(* IEC 61131-3 sources: repolevel_ST_code_completion/ground_truth/repoeval_modbus/readful_result, 6 files *)

(* ---- DataReverse_cmdReverse.st ---- *)
It seems like you are sharing code fragments from a repository, and you are particularly interested in the `cmdReverse` function and its context. However, the code snippet you provided at the end is incomplete. Let me help you understand the `cmdReverse` function and its purpose based on the fragments you have shared.

### `cmdReverse` Function Overview
The `cmdReverse` function is a simple function that takes an input of type `TargetDirect` and returns a `TargetDirect` value. The purpose of this function is to reverse the direction of a target. Based on the input value (`TargetDirect.extend` or `TargetDirect.retract`), it returns the opposite direction.

Here is the complete code for the `cmdReverse` function from the first fragment:

```pascal
FUNCTION cmdReverse : TargetDirect
VAR_INPUT
	input		:TargetDirect;
END_VAR

IF input = TargetDirect.extend THEN
	cmdReverse := TargetDirect.retract;
END_IF
IF input = TargetDirect.retract THEN
	cmdReverse := TargetDirect.extend;
END_IF
```

### Explanation
1. **Input Parameter**:
   - `input`: A variable of type `TargetDirect`, which presumably has two possible values: `extend` and `retract`.

2. **Logic**:
   - If the input is `TargetDirect.extend`, the function returns `TargetDirect.retract`.
   - If the input is `TargetDirect.retract`, the function returns `TargetDirect.extend`.

3. **Output**:
   - The function returns the reversed direction as a value of type `TargetDirect`.

### Usage Context
From the other fragments, it seems like this function is part of a larger system that involves Modbus communication and data handling. The `cmdReverse` function might be used in scenarios where the system needs to toggle or reverse the direction of a target, such as a motor or actuator.

For example:
- In the `localCmdHandler` method, variables like `exDirect` and `exeDirect` of type `TargetDirect` are declared. These might be used in conjunction with the `cmdReverse` function to handle commands that involve reversing directions.

### Missing Code
The last part of your message seems to repeat the `cmdReverse` function declaration but does not provide additional context or code. If you have specific questions or need further clarification, feel free to provide more details or ask!

(* ---- DataReverse_cmdReverse_1.st ---- *)
It seems like you are sharing code fragments from a repository, and you are particularly interested in the `cmdReverse` function and its context. However, the code snippet you provided at the end is incomplete. Let me help you understand the `cmdReverse` function and its purpose based on the fragments you have shared.

### `cmdReverse` Function Overview
The `cmdReverse` function is a simple function that takes an input of type `TargetDirect` and returns a `TargetDirect` value. The purpose of this function is to reverse the direction of a target. Based on the input value (`TargetDirect.extend` or `TargetDirect.retract`), it returns the opposite direction.

Here is the complete code for the `cmdReverse` function from the first fragment:

```pascal
FUNCTION cmdReverse : TargetDirect
VAR_INPUT
	input		:TargetDirect;
END_VAR

IF input = TargetDirect.extend THEN
	cmdReverse := TargetDirect.retract;
END_IF
IF input = TargetDirect.retract THEN
	cmdReverse := TargetDirect.extend;
END_IF
```

### Explanation
1. **Input Parameter**:
   - `input`: A variable of type `TargetDirect`, which presumably has two possible values: `extend` and `retract`.

2. **Logic**:
   - If the input is `TargetDirect.extend`, the function returns `TargetDirect.retract`.
   - If the input is `TargetDirect.retract`, the function returns `TargetDirect.extend`.

3. **Output**:
   - The function returns the reversed direction as a value of type `TargetDirect`.

### Usage Context
From the other fragments, it seems like this function is part of a larger system that involves Modbus communication and data handling. The `cmdReverse` function might be used in scenarios where the system needs to toggle or reverse the direction of a target, such as a motor or actuator.

For example:
- In the `localCmdHandler` method, variables like `exDirect` and `exeDirect` of type `TargetDirect` are declared. These might be used in conjunction with the `cmdReverse` function to handle commands that involve reversing directions.

### Missing Code
The last part of your message seems to repeat the `cmdReverse` function declaration but does not provide additional context or code. If you have specific questions or need further clarification, feel free to provide more details or ask!

(* ---- setButtonByDirect.st ---- *)
The provided code fragments define a function named `setButtonByDirect` in Structured Text (ST), which is commonly used in PLC programming. This function is designed to manipulate UI button variables based on input parameters such as `level`, `idx`, and `direct`.

### Function Overview:
- **Inputs:**
  - `level`: An integer indicating the type of track (1 for 地轨, 2 for 天轨).
  - `idx`: An integer representing the index of the挡板 (barrier).
  - `direct`: A variable of type `TargetDirect` that specifies the direction (`extend`, `retract`, or `stop`).

- **Purpose:**
  The function updates the state of UI button variables (`btnStop`, `btnExtend`, `btnRetract`) based on the input parameters.

### Key Observations:
1. **Parameter Validation:**
   - For `level = 1`, the function checks if `idx` is 0 or greater than 10. If this condition is true, the function exits early (`RETURN`).
   - For `level = 2`, the function checks if `idx` is greater than 10 and exits early if the condition is true.

2. **Button State Updates:**
   - Depending on the value of `direct` (`TargetDirect.extend`, `TargetDirect.retract`, or `TargetDirect.stop`), the function updates the button states (`btnStop`, `btnExtend`, `btnRetract`) for the specified `idx` in the `gUI.grd` array.

3. **Incomplete Code:**
   - The code fragments provided are incomplete. For example, the logic for `level = 2` is partially shown, and the handling of `TargetDirect.extend` for `level = 2` is missing.

### Suggestions for Improvement:
1. **Complete the Logic for `level = 2`:**
   - Ensure that all cases for `direct` (`extend`, `retract`, `stop`) are handled for `level = 2`.

2. **Add Comments for Clarity:**
   - While the code includes some comments, additional explanations for the logic (e.g., why certain conditions are checked) would improve readability.

3. **Error Handling:**
   - Consider adding error handling or logging for invalid input values to make debugging easier.

4. **Code Duplication:**
   - The logic for updating button states (`btnStop`, `btnExtend`, `btnRetract`) is duplicated for `level = 1` and `level = 2`. This could be refactored into a helper function to reduce redundancy.

### Example of Refactored Code:
```st
FUNCTION setButtonByDirect : BOOL
VAR_INPUT
	level		:INT;	// 1->地轨, 2->天轨
	idx			:INT;	// 挡板索引编号
	direct		:TargetDirect; // Direction
END_VAR
VAR
END_VAR

// Helper function to update button states
FUNCTION UpdateButtonStates : VOID
VAR_INPUT
	idx			:INT;
	direct		:TargetDirect;
END_VAR
BEGIN
	CASE direct OF
		TargetDirect.extend:
			gUI.grd[idx].btnStop := FALSE;
			gUI.grd[idx].btnExtend := TRUE;
			gUI.grd[idx].btnRetract := FALSE;
		TargetDirect.retract:
			gUI.grd[idx].btnStop := FALSE;
			gUI.grd[idx].btnExtend := FALSE;
			gUI.grd[idx].btnRetract := TRUE;
		TargetDirect.stop:
			gUI.grd[idx].btnStop := FALSE;
			gUI.grd[idx].btnExtend := FALSE;
			gUI.grd[idx].btnRetract := FALSE;
	END_CASE
END_FUNCTION

// Main function logic
BEGIN
	CASE level OF
		1:
			IF idx = 0 OR idx > 10 THEN
				RETURN;
			END_IF
			UpdateButtonStates(idx, direct);
		2:
			IF idx > 10 THEN
				RETURN;
			END_IF
			UpdateButtonStates(idx, direct);
	END_CASE
END_FUNCTION
```

This refactored version introduces a helper function `UpdateButtonStates` to handle button state updates, reducing code duplication and improving maintainability.

(* ---- setButtonByDirect_1.st ---- *)
The provided code fragments define a function named `setButtonByDirect` in Structured Text (ST), which is commonly used in PLC programming. This function is designed to manipulate UI button variables based on input parameters such as `level`, `idx`, and `direct`.

### Function Overview:
- **Inputs:**
  - `level`: An integer indicating the type of track (1 for 地轨, 2 for 天轨).
  - `idx`: An integer representing the index of the挡板 (barrier).
  - `direct`: A variable of type `TargetDirect` that specifies the direction (`extend`, `retract`, or `stop`).

- **Purpose:**
  The function updates the state of UI button variables (`btnStop`, `btnExtend`, `btnRetract`) based on the input parameters.

### Key Observations:
1. **Parameter Validation:**
   - For `level = 1`, the function checks if `idx` is 0 or greater than 10. If this condition is true, the function exits early (`RETURN`).
   - For `level = 2`, the function checks if `idx` is greater than 10 and exits early if the condition is true.

2. **Button State Updates:**
   - Depending on the value of `direct` (`TargetDirect.extend`, `TargetDirect.retract`, or `TargetDirect.stop`), the function updates the button states (`btnStop`, `btnExtend`, `btnRetract`) for the specified `idx` in the `gUI.grd` array.

3. **Incomplete Code:**
   - The code fragments provided are incomplete. For example, the logic for `level = 2` is partially shown, and the handling of `TargetDirect.extend` for `level = 2` is missing.

### Suggestions for Improvement:
1. **Complete the Logic for `level = 2`:**
   - Ensure that all cases for `direct` (`extend`, `retract`, `stop`) are handled for `level = 2`.

2. **Add Comments for Clarity:**
   - While the code includes some comments, additional explanations for the logic (e.g., why certain conditions are checked) would improve readability.

3. **Error Handling:**
   - Consider adding error handling or logging for invalid input values to make debugging easier.

4. **Code Duplication:**
   - The logic for updating button states (`btnStop`, `btnExtend`, `btnRetract`) is duplicated for `level = 1` and `level = 2`. This could be refactored into a helper function to reduce redundancy.

### Example of Refactored Code:
```st
FUNCTION setButtonByDirect : BOOL
VAR_INPUT
	level		:INT;	// 1->地轨, 2->天轨
	idx			:INT;	// 挡板索引编号
	direct		:TargetDirect; // Direction
END_VAR
VAR
END_VAR

// Helper function to update button states
FUNCTION UpdateButtonStates : VOID
VAR_INPUT
	idx			:INT;
	direct		:TargetDirect;
END_VAR
BEGIN
	CASE direct OF
		TargetDirect.extend:
			gUI.grd[idx].btnStop := FALSE;
			gUI.grd[idx].btnExtend := TRUE;
			gUI.grd[idx].btnRetract := FALSE;
		TargetDirect.retract:
			gUI.grd[idx].btnStop := FALSE;
			gUI.grd[idx].btnExtend := FALSE;
			gUI.grd[idx].btnRetract := TRUE;
		TargetDirect.stop:
			gUI.grd[idx].btnStop := FALSE;
			gUI.grd[idx].btnExtend := FALSE;
			gUI.grd[idx].btnRetract := FALSE;
	END_CASE
END_FUNCTION

// Main function logic
BEGIN
	CASE level OF
		1:
			IF idx = 0 OR idx > 10 THEN
				RETURN;
			END_IF
			UpdateButtonStates(idx, direct);
		2:
			IF idx > 10 THEN
				RETURN;
			END_IF
			UpdateButtonStates(idx, direct);
	END_CASE
END_FUNCTION
```

This refactored version introduces a helper function `UpdateButtonStates` to handle button state updates, reducing code duplication and improving maintainability.

(* ---- mdbsNumToIdx.st ---- *)
It seems like you are sharing multiple versions of a code fragment for a function block named `mdbsNumToIdx`. This function block takes a `devNo` (device number) as input and outputs `level` and `idx` based on the value of `devNo`. The code appears to be evolving across the fragments, with additional cases being added in each version.

Here’s a summary of the functionality and changes across the fragments:

---

### **Functionality**
1. **Input**:
   - `devNo`: A `WORD` (16-bit unsigned integer) representing the device number.

2. **Output**:
   - `level`: An `INT` (integer) representing the level associated with the device number.
   - `idx`: An `INT` representing the index associated with the device number.

3. **Logic**:
   - If `devNo > 40000`, a `CASE` statement is used to map specific `devNo` values to corresponding `level` and `idx` values.
   - The mappings are hardcoded for specific device numbers.

---

### **Code Evolution**
1. **First Fragment**:
   - Contains mappings for `devNo` values in the range `41010` to `42020`.
   - All mappings are for `level = 1`.

2. **Second Fragment**:
   - Adds mappings for `devNo` values in the range `51010` to `51040`.
   - These new mappings are for `level = 2`.

3. **Third Fragment**:
   - Extends the mappings for `level = 2` to include `devNo` values up to `51070`.

---

### **Final Version**
Here’s the consolidated version of the code based on the fragments provided:

```st
FUNCTION_BLOCK mdbsNumToIdx
VAR_INPUT
	devNo		:WORD;
END_VAR
VAR_OUTPUT
	level		:INT;
	idx			:INT;
END_VAR
VAR

END_VAR

IF devNo > 40000 THEN
	CASE devNo OF
		// 地轨 (Level 1)
		41010:	level := 1;	idx := 1;
		41020:	level := 1;	idx := 3;
		41030:	level := 1;	idx := 4;
		41040:	level := 1;	idx := 5;
		41050:	level := 1;	idx := 6;
		41060:	level := 1;	idx := 8;
		41070:	level := 1;	idx := 9;
		41080:	level := 1;	idx := 10;
		42010:	level := 1;	idx := 2;
		42020:	level := 1;	idx := 7;

		// Level 2
		51010:	level := 2;	idx := 1;
		51020:	level := 2;	idx := 3;
		51030:	level := 2;	idx := 4;
		51040:	level := 2;	idx := 5;
		51050:	level := 2;	idx := 6;
		51060:	level := 2;	idx := 8;
		51070:	level := 2;	idx := 9;
	END_CASE;
END_IF;
```

---

### **Observations**
1. **Scalability**:
   - The current implementation uses hardcoded mappings, which can become difficult to maintain as the number of `devNo` values increases.
   - Consider using a data structure (e.g., an array or a dictionary) to store the mappings, making it easier to add, remove, or modify entries.

2. **Error Handling**:
   - The code does not handle cases where `devNo` is not in the specified ranges. You might want to add a default case to handle such scenarios.

3. **Comments**:
   - The comment `//地轨` (Chinese for "ground rail") suggests that the mappings are related to specific hardware or a system. Adding more descriptive comments could help future developers understand the purpose of each mapping.

---

Let me know if you need help refactoring this code or implementing additional features!

(* ---- mdbsNumToIdx_1.st ---- *)
It seems like you are sharing multiple versions of a code fragment for a function block named `mdbsNumToIdx`. This function block takes a `devNo` (device number) as input and outputs `level` and `idx` based on the value of `devNo`. The code appears to be evolving across the fragments, with additional cases being added in each version.

Here’s a summary of the functionality and changes across the fragments:

---

### **Functionality**
1. **Input**:
   - `devNo`: A `WORD` (16-bit unsigned integer) representing the device number.

2. **Output**:
   - `level`: An `INT` (integer) representing the level associated with the device number.
   - `idx`: An `INT` representing the index associated with the device number.

3. **Logic**:
   - If `devNo > 40000`, a `CASE` statement is used to map specific `devNo` values to corresponding `level` and `idx` values.
   - The mappings are hardcoded for specific device numbers.

---

### **Code Evolution**
1. **First Fragment**:
   - Contains mappings for `devNo` values in the range `41010` to `42020`.
   - All mappings are for `level = 1`.

2. **Second Fragment**:
   - Adds mappings for `devNo` values in the range `51010` to `51040`.
   - These new mappings are for `level = 2`.

3. **Third Fragment**:
   - Extends the mappings for `level = 2` to include `devNo` values up to `51070`.

---

### **Final Version**
Here’s the consolidated version of the code based on the fragments provided:

```st
FUNCTION_BLOCK mdbsNumToIdx
VAR_INPUT
	devNo		:WORD;
END_VAR
VAR_OUTPUT
	level		:INT;
	idx			:INT;
END_VAR
VAR

END_VAR

IF devNo > 40000 THEN
	CASE devNo OF
		// 地轨 (Level 1)
		41010:	level := 1;	idx := 1;
		41020:	level := 1;	idx := 3;
		41030:	level := 1;	idx := 4;
		41040:	level := 1;	idx := 5;
		41050:	level := 1;	idx := 6;
		41060:	level := 1;	idx := 8;
		41070:	level := 1;	idx := 9;
		41080:	level := 1;	idx := 10;
		42010:	level := 1;	idx := 2;
		42020:	level := 1;	idx := 7;

		// Level 2
		51010:	level := 2;	idx := 1;
		51020:	level := 2;	idx := 3;
		51030:	level := 2;	idx := 4;
		51040:	level := 2;	idx := 5;
		51050:	level := 2;	idx := 6;
		51060:	level := 2;	idx := 8;
		51070:	level := 2;	idx := 9;
	END_CASE;
END_IF;
```

---

### **Observations**
1. **Scalability**:
   - The current implementation uses hardcoded mappings, which can become difficult to maintain as the number of `devNo` values increases.
   - Consider using a data structure (e.g., an array or a dictionary) to store the mappings, making it easier to add, remove, or modify entries.

2. **Error Handling**:
   - The code does not handle cases where `devNo` is not in the specified ranges. You might want to add a default case to handle such scenarios.

3. **Comments**:
   - The comment `//地轨` (Chinese for "ground rail") suggests that the mappings are related to specific hardware or a system. Adding more descriptive comments could help future developers understand the purpose of each mapping.

---

Let me know if you need help refactoring this code or implementing additional features!
